FUNCTION f_MakeAbsPath : STRING(255)
VAR_INPUT
	GCodePath	:	STRING(255);
END_VAR
VAR
END_VAR

f_MakeAbsPath	:=	CONCAT(UserVar.GCodeBasePath, GCodePath);

END_FUNCTION

(* stored: Version 1.1.0.1, ProductVersion 3.1.4024.15
   POU f_MakeAbsPath: Id {9bde3730-b15a-4787-9981-9d255e5c877e}, SpecialFunc None *)
